(* IEC 61131-3 sources: plc-ci-toolkit/ci/tests/samples/sa_probe_src/src/POUs/FB_SaBad, 3 files *)

(* ---- FB_SaBad.decl.st ---- *)
// Назначение: зонд статанализа (намеренно плохой код)
FUNCTION_BLOCK FB_SaBad
VAR_INPUT
    iMode : INT;
    rIn : REAL;
END_VAR
VAR_OUTPUT
    iOut : INT;
    xEqual : BOOL;
END_VAR
VAR
    {attribute 'analysis' := '-33'}
    iUnusedLocal : INT;             // SA0033 подавлено атрибутом
    iUnused2 : INT;                 // SA0033: не используется
    diWide : DINT := 70000;
    F_Clamp : REAL;                 // SA0027: имя совпадает с функцией F_Clamp
END_VAR

(* ---- Check.method.decl.st ---- *)
METHOD Check : BOOL
VAR
    fbPulse : FB_Example;           // SA0167: временный экземпляр ФБ в методе
    iNeverUsed : INT;               // SA0033 в методе
END_VAR

(* ---- FB_SaBad.impl.st ---- *)
CASE iMode OF
    1: iOut := 10;
    2: iOut := 20;
END_CASE
iOut := DINT_TO_INT(diWide);
diWide := iOut;
xEqual := rIn = 1.5;
F_Clamp := rIn;
;
IF iMode > 100 THEN
    RETURN;
    iOut := 0;
END_IF
